// TIA Portal V21 export
Screen "T07_Sym"  1024x768, Number=27
  ScreenLayer 
    SymbolicIOField "P_SymIO" at 0,0 size 100x30  Mode=Output, TextList=TL_State
      ProcessValue := State
